TYPE ET_CalcExtTrajState_1 :
(
	ET_CalcExtTrajState_eWaitExecute := 0,
	ET_CalcExtTrajState_eCalcTrajPos := 5,
	ET_CalcExtTrajState_eDone := 197,
	ET_CalcExtTrajState_eError := 198,
	ET_CalcExtTrajState_eNoExecute := 199
);
END_TYPE

(* stored: Version 1.1.0.1, ProductVersion 3.1.4024.15
   DUT ET_CalcExtTrajState_1: Id {ce4c48ce-b066-446d-a925-7ed052fd9872} *)
